# EPICS autosave request: iocBoot/iocUSB3105/auto_settings.req
file "USB3105_settings.req", P=$(P)
